(* PLC project PR_LoadingSeq_Soft2.0 1_workflow_95d36b_PLC, SiemensToBackhoff Siemens TIA Portal → Beckhoff TwinCAT PLCopen Converter 2.2 *)
(* stored: creationDateTime 2026-10-12T09:25:00.898361, modificationDateTime 2026-10-12T09:25:00.898361 *)

FUNCTION_BLOCK PR_LoadingSeq_Soft2.0 1_workflow_95d36b
VAR_INPUT
	iAbort : BOOL;
	iAcceptPartPresent : BOOL;
	iAutoRunning : BOOL;
	iFaultReset : BOOL;
	iLoadGantrySafe : BOOL;
	iOTS_Frm_Prev : BOOL;
	iPartPresent : BOOL;
	iPartPresentInGrip : BOOL;
	iRFWriteDone : BOOL;
	iRFWriteError : BOOL;
	iReject : BOOL;
	iReset_fault : BOOL;
	iRetry : BOOL;
	iRetryCount : INT;
	iSstMode : BOOL;
	iSstPB : BOOL;
	iStartFrmFibroseq : BOOL;
END_VAR
VAR_OUTPUT
	qError : ARRAY[0..1] OF BOOL;
	qLoadingOver : BOOL;
	qMessage : ARRAY[0..1] OF BOOL;
	qRTR_To_Prev : BOOL;
END_VAR
VAR
	c121_WaitForRFIDWriteOver_T1 : BOOL;
	c121_WaitForRFIDWriteOver_T2 : BOOL;
	c122_CheckRetryCountOver_T1 : BOOL;
	c122_CheckRetryCountOver_T2 : BOOL;
	c123_WaitForOperatorDecision_T1 : BOOL;
	c123_WaitForOperatorDecision_T2 : BOOL;
	c20_CheckRecoveryStatus_T1 : BOOL;
	c20_CheckRecoveryStatus_T2 : BOOL;
	c20_CheckRecoveryStatus_T3 : BOOL;
	c50_CheckPartPresentAtStation_T1 : BOOL;
	c50_CheckPartPresentAtStation_T2 : BOOL;
	c90_ConfirmPartLoad_T1 : BOOL;
	c90_ConfirmPartLoad_T2 : BOOL;
	StateNo : INT;
	s100_WaitForOperatorDecision : BOOL;
	s100_WaitForOperatorDecision_T1 : BOOL;
	s100_WaitForOperatorDecision_T2 : BOOL;
	s10_WaitForStartFrmFibroMainSeq : BOOL;
	s10_WaitForStartFrmFibroMainSeq_T1 : BOOL;
	s120_WaitForGantrySafe : BOOL;
	s120_WaitForGantrySafe_T1 : BOOL;
	s121_WaitForRFIDWriteOver : BOOL;
	s121_WaitForRFIDWriteOver_T1 : BOOL;
	s121_WaitForRFIDWriteOver_T2 : BOOL;
	s122_CheckRetryCountOver : BOOL;
	s122_CheckRetryCountOver_T1 : BOOL;
	s122_CheckRetryCountOver_T2 : BOOL;
	s123_WaitForOperatorDecision : BOOL;
	s123_WaitForOperatorDecision_T1 : BOOL;
	s123_WaitForOperatorDecision_T2 : BOOL;
	s130_WaitForStartLow : BOOL;
	s130_WaitForStartLow_T1 : BOOL;
	s1_WaitForResetRelease : BOOL;
	s1_WaitForResetRelease_T1 : BOOL;
	s20_CheckRecoveryStatus : BOOL;
	s20_CheckRecoveryStatus_T1 : BOOL;
	s20_CheckRecoveryStatus_T2 : BOOL;
	s20_CheckRecoveryStatus_T3 : BOOL;
	s30_WaitForOperatorAck : BOOL;
	s30_WaitForOperatorAck_T1 : BOOL;
	s40_WaitForLoadingGantrySafe : BOOL;
	s40_WaitForLoadingGantrySafe_T1 : BOOL;
	s50_CheckPartPresentAtStation : BOOL;
	s50_CheckPartPresentAtStation_T1 : BOOL;
	s50_CheckPartPresentAtStation_T2 : BOOL;
	s60_WaitForPartAbsentAndAck : BOOL;
	s60_WaitForPartAbsentAndAck_T1 : BOOL;
	s70_WaitForOTSFromGantry : BOOL;
	s70_WaitForOTSFromGantry_T1 : BOOL;
	s80_WaitForPartLoad : BOOL;
	s80_WaitForPartLoad_T1 : BOOL;
	s90_ConfirmPartLoad : BOOL;
	s90_ConfirmPartLoad_T1 : BOOL;
	s90_ConfirmPartLoad_T2 : BOOL;
	sAbnormalStatus : BOOL;
	sLoadInProgress : BOOL;
	sLoadInProgressInternal : INT;
	sPartPresent : BOOL;
	sRFWriteRetryCount : INT;
	sSst : BOOL;
	sSstPulse : BOOL;
	sSstRise : R_TRIG;
	sStWtResetRel : BOOL;
	sStWtResetRel_T1 : BOOL;
END_VAR
VAR_TEMP
	tOne : BOOL;
END_VAR
  VAR  (* added by the conversion: wires and edge detectors of the diagram *)
    _w24 : BOOL;
    _w26 : BOOL;
    _w39 : BOOL;
    _w41 : BOOL;
    _w42 : BOOL;
    _w59 : BOOL;
    _w62 : BOOL;
    _w63 : BOOL;
    _w96 : BOOL;
    _w99 : BOOL;
    _w100 : BOOL;
    _w101 : BOOL;
    _w102 : BOOL;
    _w115 : BOOL;
    _w117 : BOOL;
    _w118 : BOOL;
    _w135 : BOOL;
    _w137 : BOOL;
    _w138 : BOOL;
    _w162 : BOOL;
    _w164 : BOOL;
    _w165 : BOOL;
    _w166 : BOOL;
    _w180 : BOOL;
    _w182 : BOOL;
    _w183 : BOOL;
    _w196 : BOOL;
    _w200 : BOOL;
    _w201 : BOOL;
    _w219 : BOOL;
    _w222 : BOOL;
    _w223 : BOOL;
    _w254 : BOOL;
    _w256 : BOOL;
    _w257 : BOOL;
    _w258 : BOOL;
    _w274 : BOOL;
    _w276 : BOOL;
    _w277 : BOOL;
    _w278 : BOOL;
    _w295 : BOOL;
    _w298 : BOOL;
    _w299 : BOOL;
    _w323 : BOOL;
    _w327 : BOOL;
    _w328 : BOOL;
    _w329 : BOOL;
    _w367 : BOOL;
    _w369 : BOOL;
    _w370 : BOOL;
    _w371 : BOOL;
    _w400 : BOOL;
    _w402 : BOOL;
    _w403 : BOOL;
    _w404 : BOOL;
    _w429 : BOOL;
    _w432 : BOOL;
    _w433 : BOOL;
  END_VAR

(* LD diagram, written out as Structured Text *)
(* Network 1 *)
(* Create Single Step Pulse bit *)
(* Create Single Step bit *)
(* Transition for STATE Num:0 Reset Released *)
(* STATE Num:0 Reset Released *)
(* Transition for STATE Num:1 Wait For Reset Release *)
(* STATE Num:1 Wait For Reset Release *)
(* Transition for STATE Num:10 Wait For Start From Fibro Main Seq *)
(* STATE Num:10 Wait For Start From Fibro Main Seq *)
(* Condition1 for STATE Num:20 Check Recovery Status *)
(* Condition2 for STATE Num:20 Check Recovery Status *)
(* Condition3 for STATE Num:20 Check Recovery Status *)
(* Transition for STATE Num:20 Check Recovery Status *)
(* STATE Num:20 Check Recovery Status *)
(* Transition for STATE Num:30 Wait For Operator Ack *)
(* STATE Num:30 Wait For Operator Ack *)
(* Actions for STATE Num:30 Wait For Operator Ack *)
(* Transition for STATE Num:40 Wait for Loading Gantry safe *)
(* STATE Num:40 Wait for Loading Gantry safe *)
(* Condition1 for STATE Num:50 Check Part Present At Station *)
(* Condition2 for STATE Num:50 Check Part Present At Station *)
(* Transition for STATE Num:50 Check Part Present At Station *)
(* STATE Num:50 Check Part Present At Station *)
(* Transition for STATE Num:60 Wait for Part Absent And Ack *)
(* STATE Num:60 Wait for Part Absent And Ack *)
(* Transition for STATE Num:70 Wait For OTS From Gantry *)
(* STATE Num:70 Wait For OTS From Gantry *)
(* Actions for STATE Num:70 Wait For OTS From Gantry *)
(* Transition for STATE Num:80 Wait For part Load *)
(* STATE Num:80 Wait For part Load *)
(* Actions for STATE Num:80 Wait For part Load *)
(* Condition1 for STATE Num:90 Confirm Part Load *)
(* Condition2 for STATE Num:90 Confirm Part Load *)
(* Transition for STATE Num:90 Confirm Part Load *)
(* STATE Num:90 Confirm Part Load *)
(* Transition for STATE Num:100 Wait for Operator Decision *)
(* STATE Num:100 Wait for Operator Decision *)
(* Actions for STATE Num:100 Wait for Operator Decision *)
(* Transition for STATE Num:120 Wait For Gantry Safe *)
(* STATE Num:120 Wait For Gantry Safe *)
(* Condition1 for STATE Num:121 Wait For RFID Write Over *)
(* Condition2 for STATE Num:121 Wait For RFID Write Over *)
(* Transition for STATE Num:121 Wait For RFID Write Over *)
(* STATE Num:121 Wait For RFID Write Over *)
(* Actions on Transition T1 for STATE Num:121 Wait For RFID Write Over *)
(* Actions on Transition T2 for STATE Num:121 Wait For RFID Write Over *)
(* Condition1 for STATE Num:122 Check Retry Count Over *)
(* Condition2 for STATE Num:122 Check Retry Count Over *)
(* Transition for STATE Num:122 Check Retry Count Over *)
(* STATE Num:122 Check Retry Count Over *)
(* Actions on Transition T1 for STATE Num:122 Check Retry Count Over *)
(* Condition1 for STATE Num:123 Wait For Operator Decision *)
(* Condition2 for STATE Num:123 Wait For Operator Decision *)
(* Transition for STATE Num:123 Wait For Operator Decision *)
(* STATE Num:123 Wait For Operator Decision *)
(* Actions on Transition T1 for STATE Num:123 Wait For Operator Decision *)
(* Actions on Transition T2 for STATE Num:123 Wait For Operator Decision *)
(* Transition for STATE Num:130 Wait For Start Low *)
(* STATE Num:130 Wait For Start Low *)
(* Actions for STATE Num:130 Wait For Start Low *)
tOne := tOne OR NOT tOne;
sSstRise(CLK := iSstPB);
sSstPulse := sSstRise.Q;
sSst := iSstMode AND sSstPulse OR NOT iSstMode;
sStWtResetRel_T1 := sStWtResetRel AND iAutoRunning;
_w24 := sStWtResetRel;
_w26 := (_w24 OR NOT iAutoRunning) AND NOT sStWtResetRel_T1;
sStWtResetRel := _w26;
IF _w26 THEN StateNo := 0; END_IF;
s1_WaitForResetRelease_T1 := s1_WaitForResetRelease AND NOT sStWtResetRel AND sSst AND iAutoRunning;
_w39 := s1_WaitForResetRelease;
_w41 := (_w39 OR sStWtResetRel_T1) AND NOT sStWtResetRel;
_w42 := _w41 AND NOT s1_WaitForResetRelease_T1;
s1_WaitForResetRelease := _w42;
IF _w42 THEN StateNo := 1; END_IF;
s10_WaitForStartFrmFibroMainSeq_T1 := s10_WaitForStartFrmFibroMainSeq AND NOT sStWtResetRel AND sSst AND iStartFrmFibroseq;
IF s10_WaitForStartFrmFibroMainSeq AND NOT sStWtResetRel AND sSst AND iStartFrmFibroseq THEN sLoadInProgressInternal := 0; END_IF;
IF s10_WaitForStartFrmFibroMainSeq AND NOT sStWtResetRel AND sSst AND iStartFrmFibroseq THEN sRFWriteRetryCount := 0; END_IF;
_w59 := s10_WaitForStartFrmFibroMainSeq;
_w62 := (_w59 OR s130_WaitForStartLow_T1 OR s1_WaitForResetRelease_T1) AND NOT sStWtResetRel;
_w63 := _w62 AND NOT s10_WaitForStartFrmFibroMainSeq_T1;
s10_WaitForStartFrmFibroMainSeq := _w63;
IF _w63 THEN StateNo := 10; END_IF;
c20_CheckRecoveryStatus_T1 := sAbnormalStatus;
c20_CheckRecoveryStatus_T2 := sLoadInProgress;
c20_CheckRecoveryStatus_T3 := NOT sAbnormalStatus AND NOT sLoadInProgress;
s20_CheckRecoveryStatus_T1 := s20_CheckRecoveryStatus AND NOT sStWtResetRel AND sSst AND c20_CheckRecoveryStatus_T1;
s20_CheckRecoveryStatus_T2 := s20_CheckRecoveryStatus AND NOT sStWtResetRel AND sSst AND NOT s20_CheckRecoveryStatus_T1 AND c20_CheckRecoveryStatus_T2;
s20_CheckRecoveryStatus_T3 := s20_CheckRecoveryStatus AND NOT sStWtResetRel AND sSst AND NOT s20_CheckRecoveryStatus_T1 AND NOT s20_CheckRecoveryStatus_T1 AND NOT s20_CheckRecoveryStatus_T2 AND c20_CheckRecoveryStatus_T3;
_w96 := s20_CheckRecoveryStatus;
_w99 := (_w96 OR s30_WaitForOperatorAck_T1 OR s10_WaitForStartFrmFibroMainSeq_T1) AND NOT sStWtResetRel;
_w100 := _w99 AND NOT s20_CheckRecoveryStatus_T1;
_w101 := _w100 AND NOT s20_CheckRecoveryStatus_T2;
_w102 := _w101 AND NOT s20_CheckRecoveryStatus_T3;
s20_CheckRecoveryStatus := _w102;
IF _w102 THEN StateNo := 20; END_IF;
s30_WaitForOperatorAck_T1 := s30_WaitForOperatorAck AND NOT sStWtResetRel AND sSst AND iFaultReset;
_w115 := s30_WaitForOperatorAck;
_w117 := (_w115 OR s20_CheckRecoveryStatus_T1) AND NOT sStWtResetRel;
_w118 := _w117 AND NOT s30_WaitForOperatorAck_T1;
s30_WaitForOperatorAck := _w118;
IF _w118 THEN StateNo := 30; END_IF;
qError[0] := s30_WaitForOperatorAck;
s40_WaitForLoadingGantrySafe_T1 := s40_WaitForLoadingGantrySafe AND NOT sStWtResetRel AND sSst AND iLoadGantrySafe;
_w135 := s40_WaitForLoadingGantrySafe;
_w137 := (_w135 OR s20_CheckRecoveryStatus_T3) AND NOT sStWtResetRel;
_w138 := _w137 AND NOT s40_WaitForLoadingGantrySafe_T1;
s40_WaitForLoadingGantrySafe := _w138;
IF _w138 THEN StateNo := 40; END_IF;
c50_CheckPartPresentAtStation_T1 := sPartPresent;
c50_CheckPartPresentAtStation_T2 := NOT sPartPresent;
s50_CheckPartPresentAtStation_T1 := s50_CheckPartPresentAtStation AND NOT sStWtResetRel AND sSst AND c50_CheckPartPresentAtStation_T1;
s50_CheckPartPresentAtStation_T2 := s50_CheckPartPresentAtStation AND NOT sStWtResetRel AND sSst AND NOT s50_CheckPartPresentAtStation_T1 AND c50_CheckPartPresentAtStation_T2;
_w162 := s50_CheckPartPresentAtStation;
_w164 := (_w162 OR s40_WaitForLoadingGantrySafe_T1) AND NOT sStWtResetRel;
_w165 := _w164 AND NOT s50_CheckPartPresentAtStation_T1;
_w166 := _w165 AND NOT s50_CheckPartPresentAtStation_T2;
s50_CheckPartPresentAtStation := _w166;
IF _w166 THEN StateNo := 50; END_IF;
s60_WaitForPartAbsentAndAck_T1 := s60_WaitForPartAbsentAndAck AND NOT sStWtResetRel AND sSst AND (NOT iPartPresent OR iFaultReset);
_w180 := s60_WaitForPartAbsentAndAck;
_w182 := (_w180 OR s50_CheckPartPresentAtStation_T1) AND NOT sStWtResetRel;
_w183 := _w182 AND NOT s60_WaitForPartAbsentAndAck_T1;
s60_WaitForPartAbsentAndAck := _w183;
IF _w183 THEN StateNo := 60; END_IF;
s70_WaitForOTSFromGantry_T1 := s70_WaitForOTSFromGantry AND NOT sStWtResetRel AND sSst AND iOTS_Frm_Prev;
_w196 := s70_WaitForOTSFromGantry;
_w200 := (_w196 OR s100_WaitForOperatorDecision_T2 OR s60_WaitForPartAbsentAndAck_T1 OR s50_CheckPartPresentAtStation_T2) AND NOT sStWtResetRel;
_w201 := _w200 AND NOT s70_WaitForOTSFromGantry_T1;
s70_WaitForOTSFromGantry := _w201;
IF _w201 THEN StateNo := 70; END_IF;
qRTR_To_Prev := s70_WaitForOTSFromGantry;
s80_WaitForPartLoad_T1 := s80_WaitForPartLoad AND NOT sStWtResetRel AND sSst AND sPartPresent AND iLoadGantrySafe;
_w219 := s80_WaitForPartLoad;
_w222 := (_w219 OR s20_CheckRecoveryStatus_T2 OR s70_WaitForOTSFromGantry_T1) AND NOT sStWtResetRel;
_w223 := _w222 AND NOT s80_WaitForPartLoad_T1;
s80_WaitForPartLoad := _w223;
IF _w223 THEN StateNo := 80; END_IF;
IF s80_WaitForPartLoad THEN sLoadInProgressInternal := 1; END_IF;
c90_ConfirmPartLoad_T1 := NOT sPartPresent OR iPartPresentInGrip;
c90_ConfirmPartLoad_T2 := sPartPresent AND NOT iPartPresentInGrip;
s90_ConfirmPartLoad_T1 := s90_ConfirmPartLoad AND NOT sStWtResetRel AND sSst AND c90_ConfirmPartLoad_T1;
s90_ConfirmPartLoad_T2 := s90_ConfirmPartLoad AND NOT sStWtResetRel AND sSst AND NOT s90_ConfirmPartLoad_T1 AND c90_ConfirmPartLoad_T2;
_w254 := s90_ConfirmPartLoad;
_w256 := (_w254 OR s80_WaitForPartLoad_T1) AND NOT sStWtResetRel;
_w257 := _w256 AND NOT s90_ConfirmPartLoad_T1;
_w258 := _w257 AND NOT s90_ConfirmPartLoad_T2;
s90_ConfirmPartLoad := _w258;
IF _w258 THEN StateNo := 90; END_IF;
s100_WaitForOperatorDecision_T1 := s100_WaitForOperatorDecision AND NOT sStWtResetRel AND sSst AND iAcceptPartPresent;
s100_WaitForOperatorDecision_T2 := s100_WaitForOperatorDecision AND NOT sStWtResetRel AND sSst AND NOT s100_WaitForOperatorDecision_T1 AND iRetry;
_w274 := s100_WaitForOperatorDecision;
_w276 := (_w274 OR s90_ConfirmPartLoad_T1) AND NOT sStWtResetRel;
_w277 := _w276 AND NOT s100_WaitForOperatorDecision_T1;
_w278 := _w277 AND NOT s100_WaitForOperatorDecision_T2;
s100_WaitForOperatorDecision := _w278;
IF _w278 THEN StateNo := 100; END_IF;
qMessage[0] := s100_WaitForOperatorDecision;
s120_WaitForGantrySafe_T1 := s120_WaitForGantrySafe AND NOT sStWtResetRel AND sSst AND iLoadGantrySafe;
_w295 := s120_WaitForGantrySafe;
_w298 := (_w295 OR s100_WaitForOperatorDecision_T1 OR s90_ConfirmPartLoad_T2) AND NOT sStWtResetRel;
_w299 := _w298 AND NOT s120_WaitForGantrySafe_T1;
s120_WaitForGantrySafe := _w299;
IF _w299 THEN StateNo := 120; END_IF;
c121_WaitForRFIDWriteOver_T1 := iRFWriteError;
c121_WaitForRFIDWriteOver_T2 := iRFWriteDone;
s121_WaitForRFIDWriteOver_T1 := s121_WaitForRFIDWriteOver AND NOT sStWtResetRel AND sSst AND c121_WaitForRFIDWriteOver_T1;
s121_WaitForRFIDWriteOver_T2 := s121_WaitForRFIDWriteOver AND NOT sStWtResetRel AND sSst AND NOT s121_WaitForRFIDWriteOver_T1 AND c121_WaitForRFIDWriteOver_T2;
_w323 := s121_WaitForRFIDWriteOver;
_w327 := (_w323 OR s123_WaitForOperatorDecision_T2 OR s122_CheckRetryCountOver_T2 OR s120_WaitForGantrySafe_T1) AND NOT sStWtResetRel;
_w328 := _w327 AND NOT s121_WaitForRFIDWriteOver_T1;
_w329 := _w328 AND NOT s121_WaitForRFIDWriteOver_T2;
s121_WaitForRFIDWriteOver := _w329;
IF _w329 THEN StateNo := 121; END_IF;
IF s121_WaitForRFIDWriteOver_T1 THEN sRFWriteRetryCount := sRFWriteRetryCount + 1; END_IF;
qMessage[1] := s121_WaitForRFIDWriteOver_T2;
c122_CheckRetryCountOver_T1 := sRFWriteRetryCount > iRetryCount;
c122_CheckRetryCountOver_T2 := sRFWriteRetryCount <= iRetryCount;
s122_CheckRetryCountOver_T1 := s122_CheckRetryCountOver AND NOT sStWtResetRel AND sSst AND c122_CheckRetryCountOver_T1;
s122_CheckRetryCountOver_T2 := s122_CheckRetryCountOver AND NOT sStWtResetRel AND sSst AND NOT s122_CheckRetryCountOver_T1 AND c122_CheckRetryCountOver_T2;
_w367 := s122_CheckRetryCountOver;
_w369 := (_w367 OR s121_WaitForRFIDWriteOver_T1) AND NOT sStWtResetRel;
_w370 := _w369 AND NOT s122_CheckRetryCountOver_T1;
_w371 := _w370 AND NOT s122_CheckRetryCountOver_T2;
s122_CheckRetryCountOver := _w371;
IF _w371 THEN StateNo := 122; END_IF;
qError[1] := s122_CheckRetryCountOver_T1;
c123_WaitForOperatorDecision_T1 := iReject OR iAbort;
c123_WaitForOperatorDecision_T2 := iRetry;
s123_WaitForOperatorDecision_T1 := s123_WaitForOperatorDecision AND NOT sStWtResetRel AND sSst AND c123_WaitForOperatorDecision_T1;
s123_WaitForOperatorDecision_T2 := s123_WaitForOperatorDecision AND NOT sStWtResetRel AND sSst AND NOT s123_WaitForOperatorDecision_T1 AND c123_WaitForOperatorDecision_T2;
_w400 := s123_WaitForOperatorDecision;
_w402 := (_w400 OR s122_CheckRetryCountOver_T1) AND NOT sStWtResetRel;
_w403 := _w402 AND NOT s123_WaitForOperatorDecision_T1;
_w404 := _w403 AND NOT s123_WaitForOperatorDecision_T2;
s123_WaitForOperatorDecision := _w404;
IF _w404 THEN StateNo := 123; END_IF;
qMessage[1] := s123_WaitForOperatorDecision_T1;
qMessage[1] := s123_WaitForOperatorDecision_T2;
s130_WaitForStartLow_T1 := s130_WaitForStartLow AND NOT sStWtResetRel AND sSst AND NOT iStartFrmFibroseq;
IF s130_WaitForStartLow AND NOT sStWtResetRel AND sSst AND NOT iStartFrmFibroseq THEN sLoadInProgressInternal := 0; END_IF;
IF s130_WaitForStartLow AND NOT sStWtResetRel AND sSst AND NOT iStartFrmFibroseq THEN sRFWriteRetryCount := 0; END_IF;
_w429 := s130_WaitForStartLow;
_w432 := (_w429 OR s123_WaitForOperatorDecision_T1 OR s121_WaitForRFIDWriteOver_T2) AND NOT sStWtResetRel;
_w433 := _w432 AND NOT s130_WaitForStartLow_T1;
s130_WaitForStartLow := _w433;
IF _w433 THEN StateNo := 130; END_IF;
qLoadingOver := s130_WaitForStartLow;
END_FUNCTION_BLOCK
